Fanuc KAREL source: kd00038.KL

-- PROVISIONAL review KL for V770-1; original PC SHA256 e33d117685ead8fb5d3742902ae868e7f8cc2e9878afa064fd4b76149ae353ca
-- Incomplete behavior may be omitted. Consult companion uncertainty JSON. Do not deploy.
PROGRAM KD00038
%NOLOCKGROUP
VAR
  I : INTEGER
  J : INTEGER
  B : BOOLEAN
  R : REAL
  S : STRING[80]
BEGIN
  -- UNRESOLVED_PC offsets 5-18; opcodes 9D,81,18,9D,1B,9D,12,9D,13,04
  -- UNRESOLVED_PC offsets 23-27; opcodes 7F
END KD00038
